(* IEC 61131-3 sources: volt/packages/volt-lsp-iec/test-corpus/pro2193/Device/Plc Logic/Application/09 Misc/Library Manager/L_MC2P_MotionControlCam (part 2) *)

(* ---- L_MC2P_TAPPETREFTOFILE.pou ---- *)
FUNCTION_BLOCK L_MC2P_TAPPETREFTOFILE EXTENDS L_MC2P_WriteLMDFile
VAR_INPUT
	XEXECUTE : BOOL;
	SFILENAME : STRING := '';
	ITFTAPPETTABLE : L_MC2P_Tappet_REF;
END_VAR
VAR_OUTPUT
	XDONE : BOOL;
	XBUSY : BOOL;
	XERROR : BOOL;
	EERRORID : L_IE1P_Error;
END_VAR
VAR
	XRELOADOLD : BOOL;
	RELOAD : BOOL;
END_VAR
END_FUNCTION_BLOCK

METHOD MAIN
END_METHOD

METHOD WRITESPECIFICDATA
VAR_INPUT
	HFILE : SYSFILE.RTS_IEC_HANDLE;
END_VAR
END_METHOD

METHOD WRITETAPPET
VAR_INPUT
	HFILE : SYSFILE.RTS_IEC_HANDLE;
	ITFCAMDATA : L_MC2P_ITappetData;
	DWCOUNT : DWORD;
END_VAR
END_METHOD

METHOD WRITETAPPETDATA
VAR_INPUT
	HFILE : SYSFILE.RTS_IEC_HANDLE;
END_VAR
END_METHOD

(* ---- L_MC2P_TAPPETREGISTER.pou ---- *)
FUNCTION_BLOCK L_MC2P_TAPPETREGISTER EXTENDS L_MC2P_TemplateAxis_Licence
VAR_INPUT
	XENABLE : BOOL;
	XFORCE : BOOL;
	ITFTAPPETTABLE : L_MC2P_Tappet_Ref;
	LROFFSET : LREAL;
	LRHYSTERESE : LREAL;
	LRREACTTIMEON : LREAL;
	LRREACTTIMEOFF : LREAL;
	EVALUESOURCE : MC_SOURCE;
	BYDIGITALOUTPUTSEL : BYTE := 0;
	PFASTIO_OUT : POINTER TO L_FastIO_OutRef;
	XOUTPUTSTATE : BOOL := TRUE;
	XEDGECONTROL : BOOL;
END_VAR
VAR_OUTPUT
	XSWITCH : BOOL;
	XBUSY : BOOL;
	XERROR : BOOL;
	EERRORID : L_IE1P_Error;
	BYTAPPETNO : BYTE;
	LRTIMEONRELATIVE : LREAL;
	LRTIMEOFFRELATIVE : LREAL;
END_VAR
VAR
	L_MC1P_ZERODETECT1 : L_MC1P_ZeroDetect;
	PDWABSOLUTECOUNTER : POINTER TO DWORD;
	DWDUMMYCOUNTER : DWORD;
	XMAPPINGINIT : BOOL;
	LRTIMERTICK : LREAL;
	LRTIMERTICKOFF : ARRAY [0..3] OF LREAL;
	LRTIMERPOSOFFSET : ARRAY [0..3] OF LREAL;
	LRFASTIOEXTRA : LREAL := 4.0;
	DWABSOLUTECOUNTEROLD : DWORD;
	DIMAPPINGCOUNT : DINT;
	WTIMERON : WORD;
	WTIMEROFF : WORD;
	XENABLEOLD : BOOL;
	XRESETOUTPUT : BOOL;
	SCDATAOBJECT_INT : ARRAY [0..L_MC2P_InternalConst.C_TAPPETS_BUFFERSIZE] OF L_MC2P_TappetDataObject;
	SCONOFF : ARRAY [0..L_MC2P_InternalConst.C_TAPPETS_BUFFERSIZE] OF L_MC2P_TappetDataObject;
	AXCAMSWITCHEDON : ARRAY [0..L_MC2P_InternalConst.C_TAPPETS_BUFFERSIZE] OF BOOL;
	AICAMSWITCHONCYCLE : ARRAY [0..L_MC2P_InternalConst.C_TAPPETS_BUFFERSIZE] OF INT;
	AXCAMSWITCHEDOFF : ARRAY [0..L_MC2P_InternalConst.C_TAPPETS_BUFFERSIZE] OF BOOL;
	AICAMSWITCHOFFCYCLE : ARRAY [0..L_MC2P_InternalConst.C_TAPPETS_BUFFERSIZE] OF INT;
	ICYCLE : INT;
	ICYCLEFAST : INT;
	PSCTAPPETDATA_INT : POINTER TO L_MC2P_TappetData;
	DWGUID_INT : DWORD;
	LROFFSET_INT : LREAL;
	LRHYTERESE_INT : LREAL;
	LRREACTTIMEON_INT : LREAL;
	LRREACTTIMEOFF_INT : LREAL;
	EVALUESOURCE_INT : MC_SOURCE;
	LRGETPOSITION : LREAL;
	LRGETPOSITIONOLD : LREAL;
	LRCYCLELENGTH : LREAL;
	LRPOSDIFF : LREAL;
	BYDIRECTION : BYTE;
	XOFFSETCHANGE : BOOL;
	LRTAPPETON_INT : ARRAY [0..L_MC2P_InternalConst.C_TAPPETS_BUFFERSIZE] OF LREAL;
	LRTAPPETOFF_INT : ARRAY [0..L_MC2P_InternalConst.C_TAPPETS_BUFFERSIZE] OF LREAL;
	XTAPPETOK : BOOL;
	LRGETPOSITIONOLDINIT : LREAL;
	BYSTEPFASTIO : BYTE;
	BYDIRECTIONSAVE : BYTE;
	XSWITCHFASTIO : BOOL;
	UDIFASTIOORDER : UDINT;
	XFASTIOORDERSTOP : BOOL;
	BYI : BYTE;
	XFORCEFASTAKTIV : BOOL;
	UDIDX1 : UDINT;
	UDISTART1 : UDINT;
	LRINTPOSOLD : LREAL;
	XORDERPAUSE : BOOL;
	BYDIRECTIONOLD : BYTE;
	BYTAPPETIMEAKTIVE : BYTE;
	LRSWITCHTIME : LREAL;
	XTIMERSTART : BOOL;
	UDIFLAGTAPPETNO : UDINT;
	WRINGBUFFERINDEX : WORD;
	LRVELRINGBUFFER : ARRAY [0..wEncFilterCycles] OF LREAL;
	LRVELFILTERBUFFERSUM : LREAL;
	LRPOSDIFFINFILT : LREAL;
	XFLAGBUFFERFULL : BOOL;
	LRPOSDIFFHYST : LREAL;
	XHYSTERESEACTIVE : BOOL;
	XFORCEACTIVE : BOOL;
	PFREEENCODERAXIS : POINTER TO _Axis_Ref_Enc;
	EENCTYPE : L_Mc1P_EncoderType;
	LRDELAYCOMPPLCCYCLES : LREAL := 0.0;
	UDIFORINIT : UDINT;
	LRSWITCHDIFFOLD : LREAL;
	RES : INT;
	XTAPPETFREE : BOOL;
	XTAPPETOKOLD : BOOL;
	XZERO : BOOL;
	XTAPPETCLOSED : BOOL;
	XINITEDGECON : BOOL;
	XSETDELAYCOMP : BOOL;
	DWSTEADYSTATEOLD : DWORD;
	XSETDELAYCOMPOLD : BOOL;
	XDIRECTIONDETECT : BOOL;
	WCOUNTCW : WORD;
	WCOUNTCCW : WORD;
	WCOUNTMAX : WORD := 10;
	EDIRECTIONTMP : L_MC2P_Direction;
	BYDIRECTIONTMP : BYTE;
	WENCFILTERCYCLES : WORD := 10;
	LRFASTIO_OFFSETTIME : LREAL := 3;
	LRVELOCITY : LREAL;
END_VAR
END_FUNCTION_BLOCK

METHOD CALCPOSTPONE : INT
VAR_INPUT
	LRDYNAMIZE : LREAL;
	LRON : LREAL;
	LROFF : LREAL;
	LRLEN : LREAL;
END_VAR
END_METHOD

METHOD CALCTAPPETPOS : BOOL
END_METHOD

METHOD CALCTAPPETTIME : BOOL
END_METHOD

METHOD CHECKINPUTDATA : BOOL
VAR_IN_OUT
	AXIS : AXIS_REF;
END_VAR
END_METHOD

METHOD CHECKINPUTSTRUCT : BOOL
VAR_IN_OUT
	AXIS : AXIS_REF;
END_VAR
END_METHOD

METHOD CLEARMEMINTERN
END_METHOD

METHOD DIRECTIONFORCE
VAR_INPUT
	WAXISSTATE : L_MC1P_AXIS_STATE;
END_VAR
END_METHOD

METHOD DIRECTIONHYST
VAR_IN_OUT
	AXIS : AXIS_REF;
END_VAR
END_METHOD

METHOD DYNAMIZE : LREAL
VAR_INPUT
	REACTTIME : LREAL;
END_VAR
END_METHOD

METHOD GETABSOLUTECOUNTER
END_METHOD

METHOD GETPOSITION : LREAL
VAR_INPUT
	EVALUESOURCE : MC_SOURCE;
END_VAR
END_METHOD

METHOD INSERTENTRYINTOFIFO : INT
VAR_INPUT
	LRTIMERTICK : LREAL;
	BSTATE : BOOL;
END_VAR
END_METHOD

METHOD READINPUTS : BOOL
VAR_IN_OUT
	AXIS : AXIS_REF;
END_VAR
END_METHOD

METHOD RESET
END_METHOD

METHOD RESET_OUTPUTSBYERROR
VAR_INPUT
	XERROR : BOOL;
END_VAR
END_METHOD

METHOD SWITCHFASTIO
VAR_INPUT
	BYDIGITALOUTPUTSEL : BYTE;
	XHYSTERESEACTIVE : BOOL;
	LRDELAYCOM : LREAL;
END_VAR
END_METHOD

METHOD SWITCHTAPPET : BOOL
VAR_INPUT
	XENABLE : BOOL;
END_VAR
END_METHOD

METHOD CHECKDYNAMIZE : BOOL
VAR_INPUT
	LRDYNAMIZE : LREAL;
END_VAR
END_METHOD

METHOD CHECKPOS : LREAL
VAR_INPUT
	LRPOS : LREAL;
END_VAR
END_METHOD

METHOD CHECKTIME : BOOL
VAR_INPUT
	LRDYNAMIZE : LREAL;
END_VAR
END_METHOD

(* ---- L_MC2P_TEMPLATE2AXES.pou ---- *)
FUNCTION_BLOCK L_MC2P_TEMPLATE2AXES
VAR_INPUT
	MASTER : L_MC1P_IAXIS_REF_MASTERVALUES;
END_VAR
VAR_IN_OUT
	SLAVE : AXIS_REF;
END_VAR
VAR
	SINSTANCESTR : STRING;
	XERROROLD : BOOL;
	WERRORIDOLD : WORD;
	DWERRORITFID : DWORD;
	ITFMASTERVALUESDUMMY : L_MC1P_AxisMasterValuesEmpty;
END_VAR
END_FUNCTION_BLOCK

METHOD FB_GETERRORITFID : DWORD
END_METHOD

METHOD FB_RESETERROR
VAR_INPUT
	XERROR : BOOL;
	WERRORID : WORD;
END_VAR
END_METHOD

METHOD FB_SETERROR
VAR_INPUT
	WERRORID : WORD := 0;
	XSETERRORSTOP : BOOL := FALSE;
END_VAR
END_METHOD

METHOD FB_INIT : BOOL
VAR_INPUT
	BINITRETAINS : BOOL;
	BINCOPYCODE : BOOL;
END_VAR
END_METHOD

(* ---- L_MC2P_TEMPLATE2AXES_LICENCE.pou ---- *)
FUNCTION_BLOCK L_MC2P_TEMPLATE2AXES_LICENCE EXTENDS L_MC2P_Template2Axes
VAR
	LICHANDLING : L_IMHP_LLMHandling;
END_VAR
END_FUNCTION_BLOCK

METHOD ACTIVATEAPPCREDIT : BOOL
VAR_INPUT
	XACTIVATE : BOOL;
END_VAR
END_METHOD

(* ---- L_MC2P_TEMPLATE3AXES.pou ---- *)
FUNCTION_BLOCK L_MC2P_TEMPLATE3AXES
VAR_IN_OUT
	MASTER1 : AXIS_REF;
	MASTER2 : AXIS_REF;
	SLAVE : AXIS_REF;
END_VAR
VAR
	SINSTANCESTR : STRING;
	XERROROLD : BOOL;
	WERRORIDOLD : WORD;
	DWERRORITFID : DWORD;
END_VAR
END_FUNCTION_BLOCK

METHOD FB_GETERRORITFID : DWORD
END_METHOD

METHOD FB_RESETERROR
VAR_INPUT
	XERROR : BOOL;
	WERRORID : WORD;
END_VAR
END_METHOD

METHOD FB_SETERROR
VAR_INPUT
	WERRORID : WORD := 0;
	XSETERRORSTOP : BOOL := FALSE;
END_VAR
END_METHOD

METHOD FB_INIT : BOOL
VAR_INPUT
	BINITRETAINS : BOOL;
	BINCOPYCODE : BOOL;
END_VAR
END_METHOD

(* ---- L_MC2P_TEMPLATE3AXES_LICENCE.pou ---- *)
FUNCTION_BLOCK L_MC2P_TEMPLATE3AXES_LICENCE EXTENDS L_MC2P_Template3Axes
VAR
	LICHANDLING : L_IMHP_LLMHandling;
END_VAR
END_FUNCTION_BLOCK

METHOD ACTIVATEAPPCREDIT : BOOL
VAR_INPUT
	XACTIVATE : BOOL;
END_VAR
END_METHOD

(* ---- L_MC2P_TEMPLATEAXIS.pou ---- *)
FUNCTION_BLOCK L_MC2P_TEMPLATEAXIS
VAR_IN_OUT
	AXIS : AXIS_REF;
END_VAR
VAR
	SINSTANCESTR : STRING;
	XERROROLD : BOOL;
	WERRORIDOLD : WORD;
	DWERRORITFID : DWORD;
END_VAR
END_FUNCTION_BLOCK

METHOD FB_GETERRORITFID : DWORD
END_METHOD

METHOD FB_RESETERROR
VAR_INPUT
	XERROR : BOOL;
	WERRORID : WORD;
END_VAR
END_METHOD

METHOD FB_SETERROR
VAR_INPUT
	WERRORID : WORD := 0;
	XSETERRORSTOP : BOOL := FALSE;
END_VAR
END_METHOD

METHOD FB_INIT : BOOL
VAR_INPUT
	BINITRETAINS : BOOL;
	BINCOPYCODE : BOOL;
END_VAR
END_METHOD

(* ---- L_MC2P_TEMPLATEAXIS_LICENCE.pou ---- *)
FUNCTION_BLOCK L_MC2P_TEMPLATEAXIS_LICENCE EXTENDS L_MC2P_TemplateAxis
VAR
	LICHANDLING : L_IMHP_LLMHandling;
END_VAR
END_FUNCTION_BLOCK

METHOD ACTIVATEAPPCREDIT : BOOL
VAR_INPUT
	XACTIVATE : BOOL;
END_VAR
END_METHOD

(* ---- L_MC2P_TEMPLATEMASTERAXIS.pou ---- *)
FUNCTION_BLOCK L_MC2P_TEMPLATEMASTERAXIS
VAR_IN_OUT
	MASTER : AXIS_REF;
END_VAR
VAR
	SINSTANCESTR : STRING;
	XERROROLD : BOOL;
	WERRORIDOLD : WORD;
	DWERRORITFID : DWORD;
END_VAR
END_FUNCTION_BLOCK

METHOD FB_GETERRORITFID : DWORD
END_METHOD

METHOD FB_RESETERROR
VAR_INPUT
	XERROR : BOOL;
	WERRORID : WORD;
END_VAR
END_METHOD

METHOD FB_SETERROR
VAR_INPUT
	WERRORID : WORD := 0;
	XSETERRORSTOP : BOOL := FALSE;
END_VAR
END_METHOD

METHOD FB_INIT : BOOL
VAR_INPUT
	BINITRETAINS : BOOL;
	BINCOPYCODE : BOOL;
END_VAR
END_METHOD

(* ---- L_MC2P_TEMPLATENOAXIS.pou ---- *)
FUNCTION_BLOCK L_MC2P_TEMPLATENOAXIS
VAR
	SINSTANCESTR : STRING;
	XERROROLD : BOOL;
	WERRORIDOLD : WORD;
END_VAR
END_FUNCTION_BLOCK

METHOD FB_INIT : BOOL
VAR_INPUT
	BINITRETAINS : BOOL;
	BINCOPYCODE : BOOL;
END_VAR
END_METHOD

(* ---- L_MC2P_TEMPLATESLAVEAXIS.pou ---- *)
FUNCTION_BLOCK L_MC2P_TEMPLATESLAVEAXIS
VAR_IN_OUT
	SLAVE : AXIS_REF;
END_VAR
VAR
	SINSTANCESTR : STRING;
	XERROROLD : BOOL;
	WERRORIDOLD : WORD;
	DWERRORITFID : DWORD;
END_VAR
END_FUNCTION_BLOCK

METHOD FB_GETERRORITFID : DWORD
END_METHOD

METHOD FB_RESETERROR
VAR_INPUT
	XERROR : BOOL;
	WERRORID : WORD;
END_VAR
END_METHOD

METHOD FB_SETERROR
VAR_INPUT
	WERRORID : WORD := 0;
	XSETERRORSTOP : BOOL := FALSE;
END_VAR
END_METHOD

METHOD FB_INIT : BOOL
VAR_INPUT
	BINITRETAINS : BOOL;
	BINCOPYCODE : BOOL;
END_VAR
END_METHOD

(* ---- L_MC2P_WRITELMDFILE.pou ---- *)
FUNCTION_BLOCK L_MC2P_WRITELMDFILE
VAR
	TEST1 : BOOL;
	TEST2 : BOOL;
	TEST3 : BOOL;
	TEST4 : BOOL;
	SFILE_INT : STRING := '';
	EDATA_INT : L_MC2P_LMData;
	PDATA_INT : POINTER TO BYTE;
	WDATAELEMENTS_INT : WORD;
	XENABLEONLINECHANGE_INT : BOOL;
	XBUSY_INT : BOOL;
	XDONE_INT : BOOL;
	XERROR_INT : BOOL;
	EERRORID_INT : L_IE1P_Error;
	XEXECUTEOLD : BOOL;
	HFILE : SYSFILE.RTS_IEC_HANDLE;
	RES : SYSFILE.RTS_IEC_RESULT;
	ID : L_MC2P_Magic;
	DWLENGTH : DWORD;
	XACTIVECRYPTING : BOOL;
	CRYPT : Crypting;
	CK : ARRAY [0..3] OF ULINT;
	CCYCLES : WORD;
	DICDATAWRITE : DINT;
	DWSTARTCDATA : DWORD;
	ABDATA : ARRAY [0..15] OF BYTE;
	DATAIDX : DWORD;
	AVAILABLEDATA : DWORD;
	XDATAWRITEDONE : BOOL;
	UDIFSIZE : UDINT;
	UDIFBYTESWRITE : UDINT;
	RELOAD : BOOL;
END_VAR
END_FUNCTION_BLOCK

METHOD CLOSECRYPTFRAME
VAR_INPUT
	HFILE : SYSFILE.RTS_IEC_HANDLE;
END_VAR
END_METHOD

METHOD MAIN
END_METHOD

METHOD OPENCRYPTFRAME
VAR_INPUT
	HFILE : SYSFILE.RTS_IEC_HANDLE;
END_VAR
END_METHOD

METHOD RESET
END_METHOD

METHOD SETDATALENGTH
VAR_INPUT
	HFILE : SYSFILE.RTS_IEC_HANDLE;
END_VAR
END_METHOD

METHOD WRITEFRAMES
VAR_INPUT
	HFILE : SYSFILE.RTS_IEC_HANDLE;
END_VAR
END_METHOD

METHOD WRITEORGA
VAR_INPUT
	HFILE : SYSFILE.RTS_IEC_HANDLE;
END_VAR
END_METHOD

METHOD WRITESPECIFICDATA
VAR_INPUT
	HFILE : SYSFILE.RTS_IEC_HANDLE;
END_VAR
END_METHOD

METHOD CALCCRC : DWORD
VAR_INPUT
	HFILE : SYSFILE.RTS_IEC_HANDLE;
	DWLENGTH : DWORD;
END_VAR
END_METHOD

METHOD CRCCHECKSUM32BITINCREMENTAL : DWORD
VAR_INPUT
	PBDATA : POINTER TO BYTE;
	DWDATASIZE : DWORD;
	DWCRC : DWORD;
END_VAR
END_METHOD

METHOD RESETWRITEDATA
END_METHOD

METHOD CWRITECHAR
VAR_INPUT
	HFILE : SYSFILE.RTS_IEC_HANDLE;
	SDATA : STRING(16);
	N : UINT;
END_VAR
END_METHOD

METHOD CWRITEF64
VAR_INPUT
	HFILE : SYSFILE.RTS_IEC_HANDLE;
	LRDATA : LREAL;
END_VAR
END_METHOD

METHOD CWRITEU16
VAR_INPUT
	HFILE : SYSFILE.RTS_IEC_HANDLE;
	WDATA : WORD;
END_VAR
END_METHOD

METHOD CWRITEU32
VAR_INPUT
	HFILE : SYSFILE.RTS_IEC_HANDLE;
	DWDATA : DWORD;
END_VAR
END_METHOD

METHOD WRITECRYPTDATA : DWORD
VAR_INPUT
	HFILE : SYSFILE.RTS_IEC_HANDLE;
	DWSIZE : DWORD;
END_VAR
VAR_IN_OUT
	DATA : L_MC2P_IntData;
END_VAR
END_METHOD

METHOD WRITE
VAR_INPUT
	HFILE : SYSFILE.RTS_IEC_HANDLE;
	PBYBUFFER : POINTER TO BYTE;
	ULSIZE : UINT;
END_VAR
VAR_OUTPUT
	UDIDATAWRITE : UDINT;
END_VAR
END_METHOD

METHOD WRITECHAR : STRING(16)
VAR_INPUT
	HFILE : SYSFILE.RTS_IEC_HANDLE;
	SDATA : STRING(16);
	N : UINT;
END_VAR
END_METHOD

METHOD WRITEF64 : LREAL
VAR_INPUT
	HFILE : SYSFILE.RTS_IEC_HANDLE;
	LRDATA : LREAL;
END_VAR
END_METHOD

METHOD WRITEU16 : WORD
VAR_INPUT
	HFILE : SYSFILE.RTS_IEC_HANDLE;
	WDATA : WORD;
END_VAR
END_METHOD

METHOD WRITEU32
VAR_INPUT
	HFILE : SYSFILE.RTS_IEC_HANDLE;
	DWDATA : DWORD;
END_VAR
END_METHOD

METHOD ABORT : UDINT
END_METHOD

METHOD EXECUTE : UDINT
END_METHOD

(* ---- MC_CAMIN.pou ---- *)
FUNCTION_BLOCK MC_CAMIN EXTENDS L_MC2P_MasterSlaveSync
VAR_INPUT
	EXECUTE : BOOL;
	CONTINUOUSUPDATE : BOOL := FALSE;
	MASTEROFFSET : LREAL := 0;
	SLAVEOFFSET : LREAL := 0;
	MASTERSCALING : LREAL := 1;
	SLAVESCALING : LREAL := 1;
	MASTERSTARTDISTANCE : LREAL;
	MASTERSYNCPOSITION : LREAL;
	STARTMODE : MC_START_MODE := MC_Start_Mode.mcAbsolute;
	MASTERVALUESOURCE : MC_SOURCE := MC_SOURCE.mcSetValue;
	CAMTABLE : MC_CAM_REF;
	BUFFERMODE : MC_BUFFER_MODE := MC_Buffer_Mode.mcAborting;
	DIRECTCHANGE : BOOL := FALSE;
	CLUTCHTIME : LREAL := 0.001;
	VELOCITYDIFF : LREAL := 3600.0;
	ACCELERATION : LREAL := 3600.0;
	DECELERATION : LREAL := 3600.0;
	JERK : LREAL := 0.0;
	SCALINGOFFSETMODE : L_MC2P_ScalingOffsetMode := L_MC2P_ScalingOffsetMode.direct;
	PERIODIC : BOOL := TRUE;
	MASTERABSOLUTE : BOOL := TRUE;
	SLAVEABSOLUTE : BOOL := TRUE;
END_VAR
VAR_OUTPUT
	INSYNC : BOOL;
	BUSY : BOOL;
	ACTIVE : BOOL;
	COMMANDABORTED : BOOL;
	ERROR : BOOL;
	ERRORID : L_IE1P_Error;
	ENDOFPROFILE : BOOL;
END_VAR
VAR
	XPERIODIC_INT : BOOL;
	XMASTERABSOLUTE_INT : BOOL;
	XSLAVEABSOLUTE_INT : BOOL;
	PSCCAMDATA : POINTER TO L_MC2P_CamData;
	L_MC2P_FLEXCAMSTATE1 : L_MC2P_FlexCamState;
	SCINPUTMASTERSOURCE : L_MC2P_AxisProfile;
	SCACTSLAVE : L_MC2P_AxisProfile;
	SCOUTPUTSLAVE : L_MC2P_AxisProfile;
	EOFFSETMODE_INT : L_MC2P_OffsetMode;
	ESCALINGMODE_INT : L_MC2P_ScalingMode;
	ECLUTCHMODE_INT : L_MC2P_ClutchMode;
	EPOSCTRLDIRECTION_INT : L_MC2P_ReverseCtrlDirection;
	LRMASTEROFFSET_INT : LREAL;
	LRSLAVEOFFSET_INT : LREAL;
	LRMASTERSCALING_INT : LREAL;
	LRSLAVESCALING_INT : LREAL;
	LRMASTERSTARTDISTANCE_INT : LREAL;
	LRMASTERSYNCPOSITION_INT : LREAL;
	ESTARTMODE_INT : MC_START_MODE;
	EMASTERVALUESOURCE_INT : MC_SOURCE;
	EMASTERVALUESOURCE_OLD : MC_SOURCE;
	SCCAMTABLE_INT : MC_CAM_REF;
	SCCAMINFO_INT : L_MC2P_CamInfo;
	ESCALINGOFFSETMODE_INT : L_MC2P_ScalingOffsetMode;
	LRVELOCITYDIFF_INT : LREAL;
	LRACCELERATION_INT : LREAL;
	LRDECELERATION_INT : LREAL;
	LRJERK_INT : LREAL;
	XDIRECTCHANGE_INT : BOOL := FALSE;
	LRCLUTCHTIME_INT : LREAL;
	DWCHANGEID : DWORD := 1;
	STARTINCURRENTPERIOD : BOOL;
END_VAR
END_FUNCTION_BLOCK

METHOD CONVERT_CLOSEMODE
END_METHOD

METHOD CONVERT_SCALINGOFFSETMODE
END_METHOD

METHOD GET_MASTERVALUES
END_METHOD

METHOD READINPUTS
VAR_INPUT
	XREADALL : BOOL;
END_VAR
VAR_IN_OUT
	AXIS : AXIS_REF;
END_VAR
END_METHOD

METHOD RESET_OUTPUTSADD
END_METHOD

METHOD RESET_OUTPUTSBYCOMMANDABORTED
END_METHOD

METHOD RESET_OUTPUTSBYERROR
END_METHOD

METHOD SYNCIN
END_METHOD

METHOD FB_INIT : BOOL
VAR_INPUT
	BINITRETAINS : BOOL;
	BINCOPYCODE : BOOL;
END_VAR
END_METHOD

(* ---- MC_CAMOUT.pou ---- *)
FUNCTION_BLOCK MC_CAMOUT EXTENDS L_MC2P_TemplateSlaveAxis
VAR_INPUT
	EXECUTE : BOOL;
END_VAR
VAR_OUTPUT
	DONE : BOOL;
	BUSY : BOOL;
	ERROR : BOOL;
	ERRORID : L_IE1P_Error;
END_VAR
VAR
	L_MC2P_CLUTCHBASIC1 : L_MC2P_ClutchBasic;
	XSUPERIMPOSED : BOOL;
	WFUNID : WORD;
	SCINPUTSLAVE : L_MC2P_AxisProfile;
	SCOUTPUTSLAVE : L_MC2P_AxisProfile;
	XEXECUTEOLD : BOOL;
	XRESETOUTPUT : BOOL;
	LRJERK : LREAL;
	XDONEINTERN : BOOL;
	XDONEFLAG : BOOL;
END_VAR
END_FUNCTION_BLOCK

METHOD GET_SLAVEJERK
END_METHOD

METHOD GET_SLAVEVALUES
END_METHOD

METHOD RESET_OUTPUTS
END_METHOD

METHOD RESET_OUTPUTSBYCOMMANDABORTED
END_METHOD

METHOD RESET_OUTPUTSBYERROR
END_METHOD

METHOD SET_SLAVEVALUES
END_METHOD

(* ---- MC_COMBINEAXES.pou ---- *)
FUNCTION_BLOCK MC_COMBINEAXES EXTENDS L_MC2P_Template3Axes_Licence
VAR_INPUT
	EXECUTE : BOOL;
	CONTINUOUSUPDATE : BOOL := FALSE;
	COMBINEMODE : MC_COMBINE_MODE := MC_COMBINE_MODE.mcAddAxes;
	GEARRATIONUMERATORM1 : INT := 1;
	GEARRATIODENOMINATORM1 : UINT := 1;
	GEARRATIONUMERATORM2 : INT := 1;
	GEARRATIODENOMINATORM2 : UINT := 1;
	MASTERVALUESOURCEM1 : MC_SOURCE := MC_SOURCE.mcSetValue;
	MASTERVALUESOURCEM2 : MC_SOURCE := MC_SOURCE.mcSetValue;
	BUFFERMODE : MC_BUFFER_MODE := MC_Buffer_Mode.mcAborting;
	VELOCITY : LREAL := 3600.0;
	ACCELERATION : LREAL := 3600.0;
	DECELERATION : LREAL := 3600.0;
	JERK : LREAL := 0.0;
END_VAR
VAR_OUTPUT
	INSYNC : BOOL;
	BUSY : BOOL;
	ACTIVE : BOOL;
	COMMANDABORTED : BOOL;
	ERROR : BOOL;
	ERRORID : L_IE1P_Error;
END_VAR
VAR
	L_MC2P_CLUTCHBASIC1 : L_MC2P_ClutchBasic;
	L_MC2P_CAMAXISCONVERTER1 : L_MC2P_CamAxisConverter;
	L_MC2P_CAMAXISCONVERTER2 : L_MC2P_CamAxisConverter;
	L_MC2P_CAMAXISCONVERTER3 : L_MC2P_CamAxisConverter;
	L_MC2P_MODIFYAXIS1 : L_MC2P_ModifyAxis;
	L_MC2P_MODIFYAXIS2 : L_MC2P_ModifyAxis;
	XSUPERIMPOSED : BOOL;
	WFUNID : WORD;
	SCINPUTMASTERSOURCE1 : L_MC2P_AxisProfile;
	SCINPUTMASTERSOURCE2 : L_MC2P_AxisProfile;
	SCACTSLAVE : L_MC2P_AxisProfile;
	SCOUTPUTSLAVE : L_MC2P_AxisProfile;
	LRSETSCALING1 : LREAL;
	LRSETSCALING2 : LREAL;
	XEXECUTEOLD : BOOL;
	XCOMMANDABORTEDOLD : BOOL;
	INSYNCOLD : BOOL;
	XRESETOUTPUT : BOOL;
	XCONTINUOUSUPDATE : BOOL;
	XUPDATEBLOCKER : BOOL;
	UIUPDATECOUNTER : UINT;
	XCLUTCHACTIVE : BOOL;
	DWINSTANCE : __XWORD;
	XBUFFERACTIVE : BOOL;
	XPREVBUFFBDONE : BOOL;
	LRPOSOLDMASTER1 : LREAL;
	LRPOSOLDMASTER2 : LREAL;
	LRPOSMODTOLIMMASTER1 : LREAL;
	LRPOSMODTOLIMMASTER2 : LREAL;
	ECOMBINEMODE_INT : MC_COMBINE_MODE;
	IGEARRATIONUMERATORM1_INT : INT;
	UIGEARRATIODENOMINATORM1_INT : UINT := 1;
	IGEARRATIONUMERATORM2_INT : INT;
	UIGEARRATIODENOMINATORM2_INT : UINT := 1;
	EMASTERVALUESOURCEM1_INT : MC_SOURCE;
	EMASTERVALUESOURCEM2_INT : MC_SOURCE;
	LRVELOCITY_INT : LREAL;
	LRACCELERATION_INT : LREAL;
	LRDECELERATION_INT : LREAL;
	LRJERK_INT : LREAL;
	EBUFFERMODE_INT : MC_BUFFER_MODE;
	XERROR_TMP1 : BOOL;
	XERROR_TMP2 : BOOL;
	XERROR_TMP3 : BOOL;
	EERRORID_TMP1 : L_IE1P_Error;
	EERRORID_TMP2 : L_IE1P_Error;
	EERRORID_TMP3 : L_IE1P_Error;
END_VAR
END_FUNCTION_BLOCK

METHOD CALC_COMBINEAXES
END_METHOD

METHOD CHECK_AXISDATA
END_METHOD

METHOD CHECK_CONTINUOUSUPDATE
END_METHOD

METHOD CHECK_FORUPDATES
END_METHOD

METHOD GET_MASTERVALUES
END_METHOD

METHOD GET_SLAVEVALUES
END_METHOD

METHOD LOAD_AXISCONVERTER
END_METHOD

METHOD POSMASTER1MODTOLIM : LREAL
END_METHOD

METHOD POSMASTER2MODTOLIM : LREAL
END_METHOD

METHOD READINPUTS
VAR_INPUT
	XREADALL : BOOL;
END_VAR
END_METHOD

METHOD RESET_OUTPUTS
END_METHOD

METHOD RESET_OUTPUTSBYCOMMANDABORTED
END_METHOD

METHOD RESET_OUTPUTSBYERROR
END_METHOD

METHOD SET_BUFFERMODE
END_METHOD

METHOD SET_SLAVEVALUES
END_METHOD

(* ---- MC_GEARIN.pou ---- *)
FUNCTION_BLOCK MC_GEARIN EXTENDS L_MC2P_MasterSlaveSync
VAR_INPUT
	EXECUTE : BOOL;
	CONTINUOUSUPDATE : BOOL := FALSE;
	RATIONUMERATOR : INT := 1;
	RATIODENOMINATOR : UINT := 1;
	MASTERVALUESOURCE : MC_SOURCE := MC_SOURCE.mcSetValue;
	ACCELERATION : LREAL := 3600.0;
	DECELERATION : LREAL := 3600.0;
	JERK : LREAL := 0.0;
	BUFFERMODE : MC_BUFFER_MODE := MC_Buffer_Mode.mcAborting;
END_VAR
VAR_OUTPUT
	INGEAR : BOOL;
	BUSY : BOOL;
	ACTIVE : BOOL;
	COMMANDABORTED : BOOL;
	ERROR : BOOL;
	ERRORID : L_IE1P_Error;
END_VAR
VAR
	L_MC2P_CLUTCHBASIC1 : L_MC2P_ClutchBasic;
	L_MC2P_MODIFYAXIS1 : L_MC2P_ModifyAxis;
	L_MC2P_AXISCONVERTER1 : L_MC2P_AxisConverterBase;
	SCINPUTMASTERSOURCE : L_MC2P_AxisProfile;
	SCINPUTMASTERSCALED : L_MC2P_AxisProfile;
	SCACTSLAVE : L_MC2P_AxisProfile;
	SCOUTPUTSLAVE : L_MC2P_AxisProfile;
	LRPOSDIFF : LREAL;
	LRSETSCALING : LREAL;
	IRATIONUMERATOR_INT : INT;
	UIRATIODENOMINATOR_INT : UINT := 1;
	EMASTERVALUESOURCE_INT : MC_SOURCE;
	LRACCELERATION_INT : LREAL;
	LRDECELERATION_INT : LREAL;
	LRJERK_INT : LREAL;
	LROFFSET : LREAL;
	_L_MC2P_MASTERCONVERTERTOSLAVELEGTH : L_MC2P_AxisConverterBase;
	_SCINPUTMASTERCONVERTERTED : L_MC2P_AxisProfile;
	_XAXISCONVERTERCONVERTERTED : BOOL;
END_VAR
END_FUNCTION_BLOCK

METHOD CALC_SLAVEVALUES
END_METHOD

METHOD GET_MASTERVALUES
END_METHOD

METHOD READINPUTS
VAR_INPUT
	XREADALL : BOOL;
END_VAR
VAR_IN_OUT
	AXIS : AXIS_REF;
END_VAR
END_METHOD

METHOD RESET_OUTPUTSADD
END_METHOD

METHOD SET_BUFFERMODE
END_METHOD

METHOD SYNCIN
END_METHOD

METHOD FB_INIT : BOOL
VAR_INPUT
	BINITRETAINS : BOOL;
	BINCOPYCODE : BOOL;
END_VAR
END_METHOD

(* ---- MC_GEARINPOS.pou ---- *)
FUNCTION_BLOCK MC_GEARINPOS EXTENDS L_MC2P_MasterSlaveSync
VAR_INPUT
	EXECUTE : BOOL;
	RATIONUMERATOR : INT := 1;
	RATIODENOMINATOR : UINT := 1;
	MASTERVALUESOURCE : MC_SOURCE := MC_SOURCE.mcSetValue;
	MASTERSYNCPOSITION : LREAL;
	SLAVESYNCPOSITION : LREAL;
	SYNCMODE : MC_SYNC_MODE;
	MASTERSTARTDISTANCE : LREAL;
	BUFFERMODE : MC_BUFFER_MODE := MC_Buffer_Mode.mcAborting;
END_VAR
VAR_OUTPUT
	STARTSYNC : BOOL;
	INSYNC : BOOL;
	BUSY : BOOL;
	ACTIVE : BOOL;
	COMMANDABORTED : BOOL;
	ERROR : BOOL;
	ERRORID : L_IE1P_Error;
END_VAR
VAR
	L_MC2P_CLUTCHBASIC1 : L_MC2P_ClutchBasic;
	L_MC2P_MODIFYAXIS1 : L_MC2P_ModifyAxis;
	L_MC2P_AXISCONVERTER1 : L_MC2P_AxisConverterBase;
	SCINPUTMASTERSOURCE : L_MC2P_AxisProfile;
	SCINPUTMASTERSCALED : L_MC2P_AxisProfile;
	SCACTSLAVE : L_MC2P_AxisProfile;
	SCENDSLAVE : L_MC2P_AxisProfile;
	SCOUTPUTSLAVE : L_MC2P_AxisProfile;
	LRPOSDIFF : LREAL;
	LRSETSCALING : LREAL;
	LRCORRECTSYNCMODEPOS : LREAL;
	LRCALCMASTERDISTANCE : LREAL;
	IRATIONUMERATOR_INT : INT;
	UIRATIODENOMINATOR_INT : UINT := 1;
	EMASTERVALUESOURCE_INT : MC_SOURCE;
	LRMASTERSYNCPOSITION_INT : LREAL;
	LRSLAVESYNCPOSITION_INT : LREAL;
	ESYNCMODE_INT : MC_SYNC_MODE;
	LRMASTERSTARTDISTANCE_INT : LREAL;
	LRVELOCITY_INT : LREAL;
	LRACCELERATION_INT : LREAL;
	LRDECELERATION_INT : LREAL;
	LRJERK_INT : LREAL;
	LROFFSET : LREAL;
	DEBUG_INPUTMASTERPOS : LREAL;
	DEBUG_LRMASTERCLUTCHPOSITION : LREAL;
	DEBUG_LRMASTERCLUTCHDISTANCE : LREAL;
	XUSEAXISDIRECTIONINT : BOOL;
	XUSEAXISDIRECTION : BOOL := TRUE;
	USEAXISDIRECTION : BOOL;
END_VAR
END_FUNCTION_BLOCK

METHOD CALC_SLAVEENDVALUES
END_METHOD

METHOD CALC_SLAVEVALUES
END_METHOD

METHOD GET_MASTERVALUES
END_METHOD

METHOD READINPUTS
VAR_INPUT
	XREADALL : BOOL;
END_VAR
VAR_IN_OUT
	AXIS : AXIS_REF;
END_VAR
END_METHOD

METHOD RESET_OUTPUTSADD
END_METHOD

METHOD SET_BUFFERMODE_TEST
END_METHOD

METHOD SYNCIN
END_METHOD

METHOD FB_INIT : BOOL
VAR_INPUT
	BINITRETAINS : BOOL;
	BINCOPYCODE : BOOL;
END_VAR
END_METHOD

(* ---- MC_GEAROUT.pou ---- *)
FUNCTION_BLOCK MC_GEAROUT EXTENDS L_MC2P_TemplateSlaveAxis
VAR_INPUT
	EXECUTE : BOOL;
END_VAR
VAR_OUTPUT
	DONE : BOOL;
	BUSY : BOOL;
	ERROR : BOOL;
	ERRORID : L_IE1P_Error;
END_VAR
VAR
	MC_CAMOUT1 : MC_CamOut;
END_VAR
END_FUNCTION_BLOCK

(* ---- MC_PHASINGABSOLUTE.pou ---- *)
FUNCTION_BLOCK MC_PHASINGABSOLUTE EXTENDS L_MC2P_Phasing
VAR_OUTPUT
	ABSOLUTEPHASESHIFT : LREAL;
END_VAR
END_FUNCTION_BLOCK

(* ---- MC_PHASINGRELATIVE.pou ---- *)
FUNCTION_BLOCK MC_PHASINGRELATIVE EXTENDS L_MC2P_Phasing
VAR_OUTPUT
	COVEREDPHASESHIFT : LREAL;
END_VAR
END_FUNCTION_BLOCK
